(* IEC 61131-3 sources: plc-iiot-stack/src/POUs/Iiot/FB_MqttClientNone, 4 files *)

(* ---- Connect.method.decl.st ---- *)
// Реализация I_MqttClient без транспорта.
METHOD Connect : BOOL
VAR_IN_OUT CONSTANT
    // lint:allow STL007 параметр VAR_IN_OUT CONSTANT — ссылка только для чтения, а не константа
    stCfg : ST_MqttBrokerCfg;
END_VAR

(* ---- Publish.method.decl.st ---- *)
// Реализация I_MqttClient без транспорта.
METHOD Publish : BOOL
VAR_INPUT
    sTopic : STRING(GVL_Const.MQTT_TOPIC_LEN);
    eQos : E_MqttQos;
    xRetain : BOOL;
END_VAR
VAR_IN_OUT CONSTANT
    // lint:allow STL007 параметр VAR_IN_OUT CONSTANT — ссылка только для чтения, а не константа
    sPayload : STRING(GVL_Const.MQTT_PAYLOAD_LEN);
END_VAR

(* ---- Receive.method.decl.st ---- *)
// Реализация I_MqttClient без транспорта.
METHOD Receive : BOOL
VAR_IN_OUT
    sTopic : STRING(GVL_Const.MQTT_TOPIC_LEN);
    sPayload : STRING(GVL_Const.MQTT_CMD_PAYLOAD_LEN);
END_VAR
VAR_OUTPUT
    xTruncated : BOOL;
    xRetained : BOOL;
END_VAR

(* ---- Subscribe.method.decl.st ---- *)
// Реализация I_MqttClient без транспорта.
METHOD Subscribe : BOOL
VAR_INPUT
    sTopicFilter : STRING(GVL_Const.MQTT_TOPIC_LEN);
    eQos : E_MqttQos;
END_VAR
